Fanuc KAREL source: kt00089.KL

-- PROVISIONAL review KL for V1013-1; original PC SHA256 450a7c9365cc687d8e1ca57de2fdf02c3fad0e7f08653b6c82a1c6fb13e2cb7d
-- Incomplete behavior may be omitted. Consult companion uncertainty JSON. Do not deploy.
PROGRAM KT00089
%NOLOCKGROUP
VAR
  I2 : INTEGER
  OUT : INTEGER
-- UNRESOLVED_DECL H1 type=002017
BEGIN
  -- UNRESOLVED_PC offsets 5-19; opcodes 2E,22,9D,33,B4
  -- UNRESOLVED_PC offsets 24-35; opcodes 2E,23
  -- UNRESOLVED_PC offsets 40-62; opcodes 22,9D,33,B3,21,54,23
  -- UNRESOLVED_PC offsets 67-71; opcodes 7F
END KT00089
